Universal Robots URScript: EdgeProg.script

def EdgeProg():
  # Global parameters:
  global speed_ms    = 0.250
  global speed_rads  = 0.750
  global accel_mss   = 1.200
  global accel_radss = 1.200
  global blend_radius_m = 0.000

  #--------------------------
  # Add any default subprograms here
  # For example, to drive a gripper as a program call:
  # def Gripper_Open():
  #   ...
  # end
  #
  # Example to drive a spray gun:
  def SprayOn(value):
    # use the value as an output:
    DO_SPRAY = 5
    if value == 0:
      set_standard_digital_out(DO_SPRAY, False)
    else:
      set_standard_digital_out(DO_SPRAY, True)
    end
  end

  # Example to synchronize 2
  def Synchronize():
    # Use the following digital output to signal the state of the robot:
    DO_SYNC = 1

    # Use the following digital input to get the state of another robot:
    DI_SYNC = 1

    if (get_standard_digital_out(DO_SYNC) == get_standard_digital_in(DI_SYNC)):
      set_standard_digital_out(DO_SYNC, not (get_standard_digital_out(DI_SYNC)))
      sleep(0.1)
      thread Thread_wait_1():
        while (True):
          sleep(0.01)
        end
      end
      if (get_standard_digital_out(DO_SYNC) != get_standard_digital_in(DI_SYNC)):
        global thread_handler_1=run Thread_wait_1()
        while (get_standard_digital_out(DO_SYNC) != get_standard_digital_in(DI_SYNC)):
          sync()
        end
        kill thread_handler_1
      end
    else:
      if (get_standard_digital_out(DO_SYNC) != get_standard_digital_in(DI_SYNC)):
        set_standard_digital_out(DO_SYNC, not (get_standard_digital_out(DO_SYNC)))
      end
    end
  end

  #
  # Example to move an external axis
  def MoveAxis(value):
    # use the value as an output:
    DO_AXIS_1 = 1
    DI_AXIS_1 = 1
    if value <= 0:
      set_standard_digital_out(DO_AXIS_1, False)

      # Wait for digital input to change state
      #while (get_standard_digital_in(DI_AXIS_1) != False):
      #  sync()
      #end
    else:
      set_standard_digital_out(DO_AXIS_1, True)

      # Wait for digital input to change state
      #while (get_standard_digital_in(DI_AXIS_1) != True):
      #  sync()
      #end
    end
  end
  #--------------------------


  # Main program:
  # Program generated by RoboDK v6.0.7 for ABB IRB 120-3/0.6 on XX/XX/XXXX 18:00:00
  # Using nominal kinematics.
  # Using Ref. Frame Edge: p[0.100500, -0.200250, 0.300125, 0.547381, -0.295318, 0.260260]
  # set_reference(p[0.100500, -0.200250, 0.300125, 0.547381, -0.295318, 0.260260])
  # Using TCP Tool Edge: p[-0.001500, 0.002250, 0.099875, -1.759988, 1.759988, 0.729011]
  set_tcp(p[-0.001500, 0.002250, 0.099875, -1.759988, 1.759988, 0.729011])
  speed_ms    = 0.1235
  speed_rads  = 0.5818
  blend_radius_m = 0.0000
  movej([-0.087266, -0.087266, 0.261799, 0.174533, 0.698132, -0.174533],1.20000,0.58177,0,0.0000)
  blend_radius_m = 0.0125
  movel(p[-0.752411, -0.079146, 0.724974, 0.207995, 1.521767, -0.485393],accel_mss,speed_ms,0,0.013)
  halt() # reimplement this function to force stop
  sleep(1.234)
  popup("A long message with "quotes", 'apostrophes' & symbols: <>[]{}()=+-*/%;#@! and more text to make it longer than eighty characters","Message",False,False,blocking=True)
  # Comment with ; semicolon
  Gripper = ON
  set_standard_digital_out(12, False)
  Pressure = True
  while (PartPresent != True):
    sync()
  end
  while (get_standard_digital_in(7) != 1):
    sync()
  end
  DoSomething(12)
  x = 1
  movej([0.349066, -0.174533, 0.349066, 0.000000, 0.523599, 0.000000],1.20000,0.58177,0,0.0000)
  # End of main program
end

EdgeProg()
